FUNCTION F_FracR_1 : REAL
(*
Function used to get fraction part of a real number.

Constructor: 		Patryk Panylo
Company:		E. Riexinger GmbH
Date:			17.07.2014
Version:			1.00

Date:			Revision:		Who:				Comment
dd.mm.yyyy		x.xx			Initials			comment

*)
VAR_INPUT
	(* Enummerations *)

	(* Variables *)
	rReal 						:REAL;			(* Input variable *)

	(* References *)

	(* Interfaces *)

	(* Instances *)

END_VAR
VAR
	(* Enummerations *)
	
	(* Variables *)
	rFloor						:REAL;

	(* References *)

	(* Interfaces *)

	(* Instances *)

END_VAR


rFloor := DINT_TO_REAL(F_FloorDN(ABS(rReal)));								(* Floor the value *)

IF rReal < 0
THEN
	F_FracR := rReal + rFloor ;								(* The fraction of the value *)

ELSE
	F_FracR := rReal - rFloor;								(* The fraction of the value *)

END_IF

END_FUNCTION

(* stored: Version 1.1.0.1, ProductVersion 3.1.4024.15
   POU F_FracR_1: Id {44147699-db0a-47e3-85b4-4fd16cdfda10}, SpecialFunc None *)
